ADAPTER EVENT_HS (* Adapter Interface *)
  (* Standard: 61499-1 *)
  (* Version 0.0, 7/2/2026 *)
  PACKAGE Main;
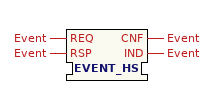
  EVENT_INPUT
    REQ; (* Request from Socket *)
    RSP; (* Response from Socket *)
  END_EVENT
  EVENT_OUTPUT
    CNF; (* Confirmation from Plug *)
    IND; (* Indication from Plug *)
  END_EVENT
  SERVICE SOCKET/PLUG
    SEQUENCE request_confirm
      SOCKET.REQ(REQD) -> PLUG.REQ(REQD);
      PLUG.CNF(CNFD) -> SOCKET.CNF(CNFD);
    END_SEQUENCE
    SEQUENCE indication_response
      PLUG.IND(INDD) -> SOCKET.IND(INDD);
      SOCKET.RSP(RSPD) -> PLUG.RSP(RSPD);
    END_SEQUENCE
  END_SERVICE
END_ADAPTER
